PROGRAM MAIN
VAR
	 // TEST ONLY - VTD MOVIPRO process data communication check.
    fbVtdProcessDataTest : FB_SEW_ProcessDataTest;
    // TEST ONLY - VTD manual control from the screen VTD_ManualTest.
    fbVtdManualControl : FB_VTD_ManualControl;
    // Safety reset from the HMI (button SAFETY RESET): one pulse per rising edge.
    rtSafetyReset : R_TRIG;
    tpSafetyReset : TP;
END_VAR

run := TRUE;

// 1. IO inputs -> internal variables
Inputs();

// 2. Logic on internal variables
// Safety reset from the HMI: one 500 ms pulse on IO_Safety.ErrorAcknowledgement and
// IO_Safety.SEW_Safety_Reset (written in Outputs). It is a request only: the TwinSAFE
// logic accepts it or not. Holding the button does not repeat the reset.
rtSafetyReset(CLK := GVL_HMI_System.stCommand.bSafetyReset);
tpSafetyReset(IN := rtSafetyReset.Q, PT := T#500MS);
Control.SafetyReset := tpSafetyReset.Q;

// TEST ONLY - two sources can write the VTD process outputs, only one at a time:
//  - the raw write of the process data screen is refused (its HMI toggle is reset)
//    while the manual screen has the drive enabled;
//  - the manual control is inhibited while the raw write is active.
IF fbVtdManualControl.q_stStatus.bEnableActive THEN
    GVL_HMI_VTD.stPdCommand.bTestWriteEnable := FALSE;
END_IF

// TEST ONLY - VTD MOVIPRO process data communication check.
fbVtdProcessDataTest(
    i_aProcessInput := Control.VTD.Motor.stProcessInput.aWord,
    i_bWcStateError := Control.VTD.Motor.stProcessInput.bWcStateError,
    i_uiEcState := Control.VTD.Motor.stProcessInput.uiEcState,
    i_bTestWriteEnable := GVL_HMI_VTD.stPdCommand.bTestWriteEnable,
    i_bTestAllowControlWord := GVL_HMI_VTD.stPdCommand.bTestAllowControlWord,
    i_aTestProcessOutput := GVL_HMI_VTD.stPdCommand.aTestProcessOutput);

// TEST ONLY - VTD manual control (jog, modes, speed, software stop, reset).
fbVtdManualControl(
    i_stProcessInput := Control.VTD.Motor.stProcessInput,
    i_bInhibit := fbVtdProcessDataTest.q_bTestWriteActive,
    i_stSettings := GVL_HMI_VTD.stManualSettings,
    io_stCommand := GVL_HMI_VTD.stManualCommand);

IF fbVtdProcessDataTest.q_bTestWriteActive THEN
    Control.VTD.Motor.aProcessOutput := fbVtdProcessDataTest.q_aProcessOutput;
ELSE
    Control.VTD.Motor.aProcessOutput := fbVtdManualControl.q_aProcessOutput;
END_IF

// 3. HMI status
FC_VTD_PdHmiUpdateStatus(
    io_fbProcessData := fbVtdProcessDataTest,
    io_stStatus := GVL_HMI_VTD.stPdStatus);
// PO really sent to the drive (raw write or manual control).
GVL_HMI_VTD.stPdStatus.aProcessOutputSent := Control.VTD.Motor.aProcessOutput;
GVL_HMI_VTD.stManualStatus := fbVtdManualControl.q_stStatus;
GVL_HMI_System.stStatus.bSafetyResetActive := tpSafetyReset.Q;

// 4. Internal variables -> IO outputs
Outputs();

END_PROGRAM

(* stored: Version 1.1.0.1
   POU MAIN: Id {324ee234-508e-4a8d-8158-a990a956945c}, SpecialFunc None *)
